(* IEC 61131-3 sources: plc-vscode/tests/st/test-ready/rusty/tests/lit/correctness/pointers/references, 4 files *)

(* ---- reference_call.st ---- *)
// RUN: (%COMPILE %s && %RUN) | %CHECK %s

FUNCTION_BLOCK fbTest
    VAR_INPUT
        reference: REF_TO BOOL; (* REF_TO *)
        p: POINTER TO BOOL;
    END_VAR
    VAR_OUTPUT
    END_VAR
    VAR_IN_OUT
        in_out1: POINTER TO BOOL; (* REF_TO *)
        in_out2: POINTER TO BOOL;
    END_VAR
    VAR
    END_VAR

    reference^ := TRUE;
    p^ := TRUE;
    in_out1^ := TRUE;
    in_out2^ := TRUE;
END_FUNCTION_BLOCK

    FUNCTION other: BOOL
    VAR
    END_VAR
    VAR_INPUT
        reference: REF_TO BOOL; (* REF_TO *)
        p: POINTER TO BOOL;
    END_VAR
    VAR_IN_OUT
        in_out1: POINTER TO BOOL; (* REF_TO *)
        in_out2: POINTER TO BOOL;
    END_VAR

    reference^ := TRUE;
    p^ := TRUE;
    in_out1^ := TRUE;
    in_out2^ := TRUE;

END_FUNCTION

FUNCTION main
VAR
    test: fbTest;
    r_a: REF_TO BOOL; (* REF_TO *)
    r_b: REF_TO BOOL; (* REF_TO *)
    p_c: POINTER TO BOOL;
    p_d: POINTER TO BOOL;
    a: BOOL := FALSE;
    b: BOOL := FALSE;
    c: BOOL := FALSE;
    d: BOOL := FALSE;
    b_result_a: BOOL := FALSE;
    b_result_b: BOOL := FALSE;
    b_result_c: BOOL := FALSE;
    b_result_d: BOOL := FALSE;
    b_result_e: BOOL := FALSE;
    b_result_f: BOOL := FALSE;
    b_result_g: BOOL := FALSE;
    b_result_h: BOOL := FALSE;
    b_result_i: BOOL := FALSE;
    b_result_j: BOOL := FALSE;
    b_result_k: BOOL := FALSE;
END_VAR
    r_a := REF(a); (* ADR *)
    p_c := r_a;
    r_a^ := TRUE;
    b_result_a := r_a^;
    b_result_b := p_c^;

    p_d := REF(d); (* ADR *)
    p_d^ := TRUE;
    b_result_c := p_d^;

    r_b := REF(b); (* ADR *)
    p_c := REF(c); (* ADR *)
    r_a^ := FALSE; r_b^ := FALSE; p_c^ := FALSE; p_d^ := FALSE;
    test(reference := r_a, p := p_c, in_out1 := r_b, in_out2 := p_d);
    b_result_d := r_a^; b_result_e := r_b^; b_result_f := p_c^; b_result_g := p_d^;

    r_a^ := FALSE; r_b^ := FALSE; p_c^ := FALSE; p_d^ := FALSE;
    other(reference := r_a, p := p_c, in_out1 := r_b, in_out2 := p_d);
    b_result_h := r_a^; b_result_i := r_b^; b_result_j := p_c^; b_result_k := p_d^;

    printf('%d$N', b_result_a); // CHECK: 1
    printf('%d$N', b_result_b); // CHECK: 1
    printf('%d$N', b_result_c); // CHECK: 1
    printf('%d$N', b_result_d); // CHECK: 1
    printf('%d$N', b_result_e); // CHECK: 1
    printf('%d$N', b_result_f); // CHECK: 1
    printf('%d$N', b_result_g); // CHECK: 1
    printf('%d$N', b_result_h); // CHECK: 1
    printf('%d$N', b_result_i); // CHECK: 1
    printf('%d$N', b_result_j); // CHECK: 1
    printf('%d$N', b_result_k); // CHECK: 1
END_FUNCTION

(* ---- reference_call_array.st ---- *)
// RUN: (%COMPILE %s && %RUN) | %CHECK %s

FUNCTION_BLOCK FbTestArray
    VAR_INPUT
        reference: REF_TO ARRAY[1..2] OF INT; (* REF_TO *)
        p: POINTER TO ARRAY[1..2] OF INT;
    END_VAR
    VAR_IN_OUT
        in_out1: REF_TO ARRAY[1..2] OF INT; (* REF_TO *)
        in_out2: POINTER TO ARRAY[1..2] OF INT;
    END_VAR

    reference^[1] := 100;
    p^[2] := 100;
    in_out1^[1] := 100;
    in_out2^[2] := 100;
END_FUNCTION_BLOCK

FUNCTION other: BOOL
    VAR_INPUT
        reference: REF_TO ARRAY[1..2] OF INT; (* REF_TO *)
        p: POINTER TO ARRAY[1..2] OF INT;
    END_VAR
    VAR_IN_OUT
        in_out1: REF_TO ARRAY[1..2] OF INT; (* REF_TO *)
        in_out2: POINTER TO ARRAY[1..2] OF INT;
    END_VAR

    reference^[1] := 100;
    p^[2] := 100;
    in_out1^[1] := 100;
    in_out2^[2] := 100;
END_FUNCTION

FUNCTION main
    VAR
        test: FbTestArray;
        a: ARRAY[1..2] OF INT;
        b: ARRAY[1..2] OF INT;
        c: ARRAY[1..2] OF INT;
        d: ARRAY[1..2] OF INT;
        ref_a: REF_TO ARRAY[1..2] OF INT; (* REF_TO *)
        ref_b: REF_TO ARRAY[1..2] OF INT; (* REF_TO *)
        p_c: POINTER TO ARRAY[1..2] OF INT;

        p_d: POINTER TO ARRAY[1..2] OF INT;
        b_result_a: INT := 0;
        b_result_b: INT := 0;
        b_result_c: INT := 0;
        b_result_d: INT := 0;
        b_result_e: INT := 0;
        b_result_f: INT := 0;
        b_result_g: INT := 0;
        b_result_h: INT := 0;
        b_result_i: INT := 0;
        b_result_j: INT := 0;
        b_result_k: INT := 0;
        b_result_l: INT := 0;
        b_result_m: INT := 0;
        b_result_n: INT := 0;
        b_result_o: INT := 0;
        b_result_p: INT := 0;
    END_VAR

        ref_a := REF(a);
        ref_b := REF(b);
        p_c := REF(c);
        p_d := REF(d);

        a[1] := 0; a[2] := 0;
        b[1] := 0; b[2] := 0;
        c[1] := 0; c[2] := 0;
        d[1] := 0; d[2] := 0;

        other(reference := ref_a, p := p_c, in_out1 := ref_b, in_out2 := p_d);
        b_result_a := a[1];
        b_result_b := a[2];
        b_result_c := b[1];
        b_result_d := b[2];
        b_result_e := c[1];
        b_result_f := c[2];
        b_result_g := d[1];
        b_result_h := d[2];

        a[1] := 0; a[2] := 0;
        b[1] := 0; b[2] := 0;
        c[1] := 0; c[2] := 0;
        d[1] := 0; d[2] := 0;

        test(reference := ref_a, p := p_c, in_out1 := ref_b, in_out2 := p_d);
        b_result_i := a[1];
        b_result_j := a[2];
        b_result_k := b[1];
        b_result_l := b[2];
        b_result_m := c[1];
        b_result_n := c[2];
        b_result_o := d[1];
        b_result_p := d[2];

    printf('%d$N', b_result_a); // CHECK: 100
    printf('%d$N', b_result_b); // CHECK: 0
    printf('%d$N', b_result_c); // CHECK: 100
    printf('%d$N', b_result_d); // CHECK: 0
    printf('%d$N', b_result_e); // CHECK: 0
    printf('%d$N', b_result_f); // CHECK: 100
    printf('%d$N', b_result_g); // CHECK: 0
    printf('%d$N', b_result_h); // CHECK: 100
    printf('%d$N', b_result_i); // CHECK: 100
    printf('%d$N', b_result_j); // CHECK: 0
    printf('%d$N', b_result_k); // CHECK: 100
    printf('%d$N', b_result_l); // CHECK: 0
    printf('%d$N', b_result_m); // CHECK: 0
    printf('%d$N', b_result_n); // CHECK: 100
    printf('%d$N', b_result_o); // CHECK: 0
    printf('%d$N', b_result_p); // CHECK: 100
END_FUNCTION

(* ---- reference_call_struct.st ---- *)
// RUN: (%COMPILE %s && %RUN) | %CHECK %s

TYPE MyStruct:
STRUCT
    field1: BOOL;
    field2: INT;
END_STRUCT
END_TYPE

FUNCTION_BLOCK FbTestStruct
    VAR_INPUT
        reference: REF_TO MyStruct; (* REF_TO *)
        p: POINTER TO MyStruct;
    END_VAR
    VAR_OUTPUT
    END_VAR
    VAR_IN_OUT
        in_out1: REF_TO MyStruct; (* REF_TO *)
        in_out2: POINTER TO MyStruct;
    END_VAR

    reference^.field1 := TRUE;
    p^.field2 := 100;
    in_out1^.field1 := TRUE;
    in_out2^.field2 := 100;
END_FUNCTION_BLOCK

FUNCTION other: BOOL
    VAR
    END_VAR
    VAR_INPUT
        reference: REF_TO MyStruct; (* REF_TO *)
        p: POINTER TO MyStruct;
    END_VAR

    VAR_IN_OUT
        in_out1: REF_TO MyStruct; (* REF_TO *)
        in_out2: POINTER TO MyStruct;
    END_VAR

    reference^.field1 := TRUE;
    p^.field2 := 100;
    in_out1^.field1 := TRUE;
    in_out2^.field2 := 100;
END_FUNCTION

FUNCTION main
    VAR
        test: FbTestStruct;
        a: MyStruct;
        b: MyStruct;
        ref_a: REF_TO MyStruct; (* REF_TO *)
        ref_b: REF_TO MyStruct; (* REF_TO *)
        p_a: POINTER TO MyStruct;
        p_b: POINTER TO MyStruct;
        b_result_a: BOOL := FALSE;
        b_result_b: INT := 0;
        b_result_c: BOOL := FALSE;
        b_result_d: INT := 0;
        b_result_e: BOOL := FALSE;
        b_result_f: INT := 0;
        b_result_g: BOOL := FALSE;
        b_result_h: INT := 0;
    END_VAR
        a.field1 := FALSE; a.field2 := 0;
        b.field1 := FALSE; b.field2 := 0;

        ref_a := REF(a);
        ref_b := REF(b);
        p_a := REF(a);
        p_b := REF(b);
        other(reference := ref_a, p := p_a, in_out1 := ref_b, in_out2 := p_b);
        b_result_a := a.field1;
        b_result_b := a.field2;
        b_result_c := b.field1;
        b_result_d := b.field2;

        a.field1 := FALSE; a.field2 := 0;
        b.field1 := FALSE; b.field2 := 0;

        test(reference := ref_a, p := ref_a, in_out1 := ref_b, in_out2 := ref_b);
        b_result_e := a.field1;
        b_result_f := a.field2;
        b_result_g := b.field1;
        b_result_h := b.field2;

    printf('%d$N', b_result_a); // CHECK: 1
    printf('%d$N', b_result_b); // CHECK: 100
    printf('%d$N', b_result_c); // CHECK: 1
    printf('%d$N', b_result_d); // CHECK: 100
    printf('%d$N', b_result_e); // CHECK: 1
    printf('%d$N', b_result_f); // CHECK: 100
    printf('%d$N', b_result_g); // CHECK: 1
    printf('%d$N', b_result_h); // CHECK: 100
END_FUNCTION

(* ---- reference_initialization.st ---- *)
// RUN: (%COMPILE %s && %RUN) | %CHECK %s

FUNCTION_BLOCK F1
VAR
    a: INT;
    b: DINT;
END_VAR
END_FUNCTION_BLOCK

PROGRAM mainProg
VAR
    myInt: INT;
    myRefInt: REF_TO INT := REF(myInt);
    myF1: F1;
    myRefF1: REF_TO F1 := REF(myF1);
END_VAR
END_PROGRAM

FUNCTION main
VAR
    tmpInt: INT;
    tmpA: INT;
    tmpB: DINT;
END_VAR
    // Initialize through direct variables
    mainProg.myInt := 11;
    mainProg.myF1.a := 22;
    mainProg.myF1.b := 33;

    // Read through references
    tmpInt := mainProg.myRefInt^;
    tmpA := mainProg.myRefF1^.a;
    tmpB := mainProg.myRefF1^.b;

    printf('ref_read_int=%d$N', tmpInt); // CHECK: ref_read_int=11
    printf('ref_read_f1_a=%d$N', tmpA); // CHECK: ref_read_f1_a=22
    printf('ref_read_f1_b=%d$N', tmpB); // CHECK: ref_read_f1_b=33

    // Write through references
    mainProg.myRefInt^ := 44;
    mainProg.myRefF1^.a := 55;
    mainProg.myRefF1^.b := 66;

    printf('direct_read_int=%d$N', mainProg.myInt); // CHECK: direct_read_int=44
    printf('direct_read_f1_a=%d$N', mainProg.myF1.a); // CHECK: direct_read_f1_a=55
    printf('direct_read_f1_b=%d$N', mainProg.myF1.b); // CHECK: direct_read_f1_b=66
END_FUNCTION
